TYPE stShutterConfig :
STRUCT
    TravelTime : TIME := T#30S;			// Time for full open/close vertical movement
	AngleFullTurnTime : TIME := T#3S;			// Time for fins to make full rotation
	TravelTimeOverstep : TIME := T#500MS;		// High state output signal time allowed to be maintain after reaching full open position
END_STRUCT
END_TYPE

(* stored: Version 1.1.0.1
   DUT stShutterConfig: Id {cba03735-b58c-4ca0-9c02-4878db374737} *)
